Staubli VAL3: readData.pgx

program readData(sio& x_UdpSocket, num& x_nData[], bool& x_bNewData, bool& x_bError)
  local bool l_bNewData
  local bool l_bError
  local num l_nMaxAttempts
  local num l_nAttempt
begin

  l_bNewData = false
  l_bError = false
  l_nMaxAttempts = 2
  l_nAttempt = 1

  // Initialize output flags
  x_bNewData = l_bNewData
  x_bError = l_bError

  // Try to read from UDP socket multiple times
  while(l_nAttempt <= l_nMaxAttempts)
    call readDataOnce(x_UdpSocket, x_nData, l_bNewData, l_bError)

    // If error, set error and exit
    if(l_bError)
      logMsg("ros2_server::readData : communication error", 2)
      x_bNewData = false
      x_bError = true
      return
    endIf

    // If new (valid) data received, set flag
    if(l_bNewData)
      // Successfully read a new message
      x_bNewData = true
    endIf

    // If data received, but last attempt did not yield new data, exit
    if(x_bNewData and !l_bNewData)
      return
    endIf

    // Prepare next attempt
    l_nAttempt = l_nAttempt + 1
  endWhile
end
